Fanuc KAREL source: kd00038.KL

-- PROVISIONAL review KL for V1013-1; original PC SHA256 3b73a98277ce5d15c394180431436d7bedb1f15aa3c4ac0a0e95d69e84fb110b
-- Incomplete behavior may be omitted. Consult companion uncertainty JSON. Do not deploy.
PROGRAM KD00038
%NOLOCKGROUP
VAR
  I : INTEGER
  J : INTEGER
  B : BOOLEAN
  R : REAL
  S : STRING[80]
BEGIN
  -- UNRESOLVED_PC offsets 5-18; opcodes 9D,81,18,9D,1B,9D,12,9D,13,04
  -- UNRESOLVED_PC offsets 23-27; opcodes 7F
END KD00038
